(* IEC 61131-3 sources: sceptre-phenix-topologies/cherrymountain-brewery/plant/generated/ci/openplc/plc-cellar, 1 file *)

(* ---- located_vars.st ---- *)
(* Generated by plantgen from plant/plant.yaml (variant ci). Do not edit. *)
(* Analog values are raw registers: engineering value = raw / 10^scaling. *)
(* RIO I/O is at %IX100.0 / %QX100.0 / %IW100 / %QW100 (v3 and v4 alike). *)
(* PLC memory: bits from %QX0.0 (coils), words from %MW0 (holding register qw_count and up, see modbus_slave.json). *)
VAR
  CEL_CLK_KI01_PV AT %IW100 : UINT; (* Cellar simulation clock (compressed fermentation time), h, x10 *)
  CEL_FV101_TT01_PV AT %IW101 : UINT; (* FV-101 side temperature, degF, x100 *)
  CEL_FV101_TT01_ALM_DEVIATION AT %QX0.0 : BOOL; (* FV-101 side temperature: deviation alarm (high) *)
  CEL_FV101_TT01_ALM_HIGH AT %QX0.1 : BOOL; (* FV-101 side temperature: high alarm (medium) *)
  CEL_FV101_TV01_CMD AT %QX100.0 : BOOL; (* FV-101 side glycol valve command *)
  CEL_FV101_TT02_PV AT %IW102 : UINT; (* FV-101 cone temperature, degF, x100 *)
  CEL_FV101_TT02_ALM_DEVIATION AT %QX0.2 : BOOL; (* FV-101 cone temperature: deviation alarm (medium) *)
  CEL_FV101_TV02_CMD AT %QX100.1 : BOOL; (* FV-101 cone glycol valve command *)
  CEL_FV101_PT01_PV AT %IW103 : UINT; (* FV-101 head pressure (absolute), psia, x100 *)
  CEL_FV101_PT01_ALM_HIGH AT %QX0.3 : BOOL; (* FV-101 head pressure (absolute): high alarm (high) *)
  CEL_FV101_PT01_ALM_LOW AT %QX0.4 : BOOL; (* FV-101 head pressure (absolute): low alarm (low) *)
  CEL_FV101_DT01_PV AT %IW104 : UINT; (* FV-101 apparent extract (sample-port density meter), degP, x100 *)
  CEL_FV101_PCV01_SP AT %QW100 : UINT; (* FV-101 spunding valve setpoint (absolute), psia, x100 *)
  CEL_FV101_ZSO01_PV AT %IX100.0 : BOOL; (* FV-101 spunding valve open (venting) *)
  CEL_FV101_TT01_SP AT %MW0 : UINT; (* FV-101 side temperature setpoint, degF, x100 *)
  CEL_FV101_TT02_SP AT %MW1 : UINT; (* FV-101 cone temperature setpoint, degF, x100 *)
  CEL_FV102_TT01_PV AT %IW105 : UINT; (* FV-102 side temperature, degF, x100 *)
  CEL_FV102_TT01_ALM_DEVIATION AT %QX0.5 : BOOL; (* FV-102 side temperature: deviation alarm (high) *)
  CEL_FV102_TT01_ALM_HIGH AT %QX0.6 : BOOL; (* FV-102 side temperature: high alarm (medium) *)
  CEL_FV102_TV01_CMD AT %QX100.2 : BOOL; (* FV-102 side glycol valve command *)
  CEL_FV102_TT02_PV AT %IW106 : UINT; (* FV-102 cone temperature, degF, x100 *)
  CEL_FV102_TT02_ALM_DEVIATION AT %QX0.7 : BOOL; (* FV-102 cone temperature: deviation alarm (medium) *)
  CEL_FV102_TV02_CMD AT %QX100.3 : BOOL; (* FV-102 cone glycol valve command *)
  CEL_FV102_PT01_PV AT %IW107 : UINT; (* FV-102 head pressure (absolute), psia, x100 *)
  CEL_FV102_PT01_ALM_HIGH AT %QX1.0 : BOOL; (* FV-102 head pressure (absolute): high alarm (high) *)
  CEL_FV102_PT01_ALM_LOW AT %QX1.1 : BOOL; (* FV-102 head pressure (absolute): low alarm (low) *)
  CEL_FV102_DT01_PV AT %IW108 : UINT; (* FV-102 apparent extract (sample-port density meter), degP, x100 *)
  CEL_FV102_PCV01_SP AT %QW101 : UINT; (* FV-102 spunding valve setpoint (absolute), psia, x100 *)
  CEL_FV102_ZSO01_PV AT %IX100.1 : BOOL; (* FV-102 spunding valve open (venting) *)
  CEL_FV102_TT01_SP AT %MW2 : UINT; (* FV-102 side temperature setpoint, degF, x100 *)
  CEL_FV102_TT02_SP AT %MW3 : UINT; (* FV-102 cone temperature setpoint, degF, x100 *)
  CEL_FV103_TT01_PV AT %IW109 : UINT; (* FV-103 side temperature, degF, x100 *)
  CEL_FV103_TT01_ALM_DEVIATION AT %QX1.2 : BOOL; (* FV-103 side temperature: deviation alarm (high) *)
  CEL_FV103_TT01_ALM_HIGH AT %QX1.3 : BOOL; (* FV-103 side temperature: high alarm (medium) *)
  CEL_FV103_TV01_CMD AT %QX100.4 : BOOL; (* FV-103 side glycol valve command *)
  CEL_FV103_TT02_PV AT %IW110 : UINT; (* FV-103 cone temperature, degF, x100 *)
  CEL_FV103_TT02_ALM_DEVIATION AT %QX1.4 : BOOL; (* FV-103 cone temperature: deviation alarm (medium) *)
  CEL_FV103_TV02_CMD AT %QX100.5 : BOOL; (* FV-103 cone glycol valve command *)
  CEL_FV103_PT01_PV AT %IW111 : UINT; (* FV-103 head pressure (absolute), psia, x100 *)
  CEL_FV103_PT01_ALM_HIGH AT %QX1.5 : BOOL; (* FV-103 head pressure (absolute): high alarm (high) *)
  CEL_FV103_PT01_ALM_LOW AT %QX1.6 : BOOL; (* FV-103 head pressure (absolute): low alarm (low) *)
  CEL_FV103_DT01_PV AT %IW112 : UINT; (* FV-103 apparent extract (sample-port density meter), degP, x100 *)
  CEL_FV103_PCV01_SP AT %QW102 : UINT; (* FV-103 spunding valve setpoint (absolute), psia, x100 *)
  CEL_FV103_ZSO01_PV AT %IX100.2 : BOOL; (* FV-103 spunding valve open (venting) *)
  CEL_FV103_TT01_SP AT %MW4 : UINT; (* FV-103 side temperature setpoint, degF, x100 *)
  CEL_FV103_TT02_SP AT %MW5 : UINT; (* FV-103 cone temperature setpoint, degF, x100 *)
  CEL_FV104_TT01_PV AT %IW113 : UINT; (* FV-104 side temperature, degF, x100 *)
  CEL_FV104_TT01_ALM_DEVIATION AT %QX1.7 : BOOL; (* FV-104 side temperature: deviation alarm (high) *)
  CEL_FV104_TT01_ALM_HIGH AT %QX2.0 : BOOL; (* FV-104 side temperature: high alarm (medium) *)
  CEL_FV104_TV01_CMD AT %QX100.6 : BOOL; (* FV-104 side glycol valve command *)
  CEL_FV104_TT02_PV AT %IW114 : UINT; (* FV-104 cone temperature, degF, x100 *)
  CEL_FV104_TT02_ALM_DEVIATION AT %QX2.1 : BOOL; (* FV-104 cone temperature: deviation alarm (medium) *)
  CEL_FV104_TV02_CMD AT %QX100.7 : BOOL; (* FV-104 cone glycol valve command *)
  CEL_FV104_PT01_PV AT %IW115 : UINT; (* FV-104 head pressure (absolute), psia, x100 *)
  CEL_FV104_PT01_ALM_HIGH AT %QX2.2 : BOOL; (* FV-104 head pressure (absolute): high alarm (high) *)
  CEL_FV104_PT01_ALM_LOW AT %QX2.3 : BOOL; (* FV-104 head pressure (absolute): low alarm (low) *)
  CEL_FV104_DT01_PV AT %IW116 : UINT; (* FV-104 apparent extract (sample-port density meter), degP, x100 *)
  CEL_FV104_PCV01_SP AT %QW103 : UINT; (* FV-104 spunding valve setpoint (absolute), psia, x100 *)
  CEL_FV104_ZSO01_PV AT %IX100.3 : BOOL; (* FV-104 spunding valve open (venting) *)
  CEL_FV104_TT01_SP AT %MW6 : UINT; (* FV-104 side temperature setpoint, degF, x100 *)
  CEL_FV104_TT02_SP AT %MW7 : UINT; (* FV-104 cone temperature setpoint, degF, x100 *)
END_VAR
